// TIA Portal V20 export
// export: Created 2026-10-20T12:52:44.0484529Z, ExportSetting WithDefaults, DisplayName Totally Integrated Automation Portal, DisplayVersion V20 Update 6, DisplayName TIA Portal Openness, DisplayVersion V20 Update 6, DisplayName TIA Portal Version Control Interface, DisplayVersion V20 Update 6, DisplayName SINAMICS Startdrive Advanced, DisplayVersion V20 SP1, DisplayName SINAMICS Startdrive G130, G150, S120, S150, SINAMICS MV, G220, S200, S210, DisplayVersion V20 SP1, DisplayName SINAMICS Startdrive G110M, G120, G120C, G120D, G120P, G115D, DisplayVersion V20 SP1, DisplayName STEP 7 Professional, DisplayVersion V20 Update 6, DisplayName STEP 7 Safety, DisplayVersion V20 Update 2, DisplayName WinCC Basic/Comfort/Advanced, DisplayVersion V20 Update 6, DisplayName WinCC Unified, DisplayVersion V20 Update 6
FUNCTION "Gate_Status_Update_FC" : Void   // FC49, SCL
{ S7_Optimized_Access := 'TRUE' }
VERSION : 0.1
// stored: AutoNumber true, IsIECCheckEnabled false, SetENOAutomatically false, UDAEnableTagReadback false
   VAR_INPUT
      Gate_Index : Int;
      Request_Access : Bool;
      Stop_Mode_Granted : Bool;
   END_VAR
   VAR_OUTPUT
      DB_SM_To_LGX_Gate_Status : Array[0..10] of Byte;
   END_VAR
   VAR_TEMP
      tGateByte : Byte;
   END_VAR
BEGIN
   #tGateByte := 0;

   IF #Request_Access THEN
       #tGateByte := #tGateByte OR BYTE#16#01;
   END_IF; // Bit 0
   IF #Stop_Mode_Granted THEN
       #tGateByte := #tGateByte OR BYTE#16#02;
   END_IF; // Bit 1
   // Bits 2..7: Free

   IF #Gate_Index >= 0 AND #Gate_Index <= 10 THEN
       #DB_SM_To_LGX_Gate_Status[#Gate_Index] := #tGateByte;
   END_IF;
END_FUNCTION
